Fanuc KAREL source: KT00809.KL

PROGRAM KT00809
%NOLOCKGROUP
VAR
  I1: INTEGER
  I2: INTEGER
  OUT: REAL
BEGIN
  I1 = 2
  I2 = 3
  I1 = 2
  I2 = 3
  OUT = LN(I1)
END KT00809
